(* IEC 61131-3 sources: nautilus/website/lessons/b4-counter/variants/ok-r-trig-then-ctu, 1 file *)

(* ---- program.st ---- *)
PROGRAM Counter
VAR edge : R_TRIG; parcels : CTU; END_VAR
edge(CLK := Eye);
parcels(CU := edge.Q, R := Reset, PV := 5);
Count := parcels.CV;
Full := parcels.Q;
END_PROGRAM
